// TIA Portal V19 export
DATA_BLOCK "R17_DATA"   // DB43
{ S7_Optimized_Access := 'FALSE' }
   VAR RETAIN
      R17 : Struct
         START : Bool;
         Reset : Bool;
         "E stop" : Bool;
         RUNNING : Bool;
         "STEP" : Int;
         START_PLS : Bool;
         STOP_PLS : Bool;
         COOL_RUNNING : Bool;
         "HEAT RUNNING" : Bool;
         TEMP_SP : Real;
         TOLERANCE_SP : Real;
         "CONTROL TYPE" : Int;
         PV : Real;
         PRODUCT_TT : Real;
         PUMP_CMD : Bool;
         TOLERANCE_MET : Bool;
         CTS_CMD : Bool;
         CTR_CMD : Bool;
         UCHWS_CMD : Bool;
         CHWS_CMD : Bool;
         HWS_CMD : Bool;
         UCHWR_CMD : Bool;
         CHWR_CMD : Bool;
         HWR_CMD : Bool;
         CTS_CMD_1 : Bool;
         CTR_CMD_1 : Bool;
         UCHWS_CMD_1 : Bool;
         CHWS_CMD_1 : Bool;
         HWS_CMD_1 : Bool;
         UCHWR_CMD_1 : Bool;
         CHWR_CMD_1 : Bool;
         HWR_CMD_1 : Bool;
         CTS_CMD_2 : Bool;
         CTR_CMD_2 : Bool;
         UCHWS_CMD_2 : Bool;
         CHWS_CMD_2 : Bool;
         HWS_CMD_2 : Bool;
         UCHWR_CMD_2 : Bool;
         CHWR_CMD_2 : Bool;
         HWR_CMD_2 : Bool;
         JACKET_CONTROL : Bool;
         RAMP_MASS : Bool;
         PRODUCT_CONTROL : Bool;
         COOL_UCH_MIN_SP : Real := 14.0;
         COOL_UCH_MAX_SP : Real := -20.0;
         COOL_CH_MIN_SP : Real := 50.0;
         COOL_CH_MAX_SP : Real := 15.0;
         COOL_CT_MIN_SP : Real := 89.0;
         COOL_CT_MAX_SP : Real := 60.0;
         COOL_HW_MIN_SP : Real := 120.0;
         COOL_HW_MAX_SP : Real := 90.0;
         HEAT_UCH_MIN_SP : Real := -20.0;
         HEAT_UCH_MAX_SP : Real := -10.0;
         HEAT_CH_MIN_SP : Real := -9.9;
         HEAT_CH_MAX_SP : Real := 5.0;
         HEAT_CT_MIN_SP : Real := 4.9;
         HEAT_CT_MAX_SP : Real := 24.0;
         HEAT_HW_MIN_SP : Real := 25.0;
         HEAT_HW_MAX_SP : Real := 120.0;
         SELECT_UCHWS : Bool;
         SELECT_CHWS : Bool;
         SELECT_CTS : Bool;
         SELECT_HWS : Bool;
         UCHWS_IN : Bool;
         CHWS_IN : Bool;
         CTS_IN : Bool;
         HWS_IN : Bool;
         UCHWS_OUT : Bool;
         CHWS_OUT : Bool;
         CTS_OUT : Bool;
         HWS_OUT : Bool;
         RAMP_START : Bool;
         RAMP_INPUT : Real;
         MAIN_TIME : Int;
         MAIN_RESET : Bool;
         RAMP_TIME : Int := 0;
         RAMP_RATE : Real;
         MAIN_COMPLETED : Bool;
         UTILITY_SEL : Int;
         REF_TT : Int;
         STEP_NO : Int;
         MAIN_PV : Real;
         CSV_CMD_3 : Bool;
         CRV_CMD_4 : Bool;
         NORM_MIN : Int;
         NORM_MAX : Int := 27684;
         NORM_OUT : Real;
         SCALE_MIN : Real;
         SCALE_MAX : Real := 100.0;
         SCVOUT : Int;
         MAN_OUT : Int;
         MAN_INPUT : Int;
         AO : Int;
         TIMER_RESET : Bool;
         COOL_CHWS_CMD : Bool;
         COOL_PUMP_CMD : Bool;
         COOL_CV_CMD : Bool;
         COOL_CS_CMD : Bool;
         COOL_HS_CMD : Bool;
         COOL_UCHS_CMD : Bool;
         R17_ramp_substitute : Real;
         COL_UTILITY_SEL : Int;
         HET_UTILITY_SEL : Int;
         AO_REVERSE : Int;
         RAMP_TMR : Int;
      END_STRUCT;
   END_VAR
BEGIN
END_DATA_BLOCK
